Fanuc KAREL source: KT00808.KL

PROGRAM KT00808
%NOLOCKGROUP
VAR
  I1: INTEGER
  I2: INTEGER
  OUT: INTEGER
BEGIN
  I1 = 2
  I2 = 3
  I1 = 2
  I2 = 3
  OUT = LN(I1)
END KT00808
